Fanuc KAREL source: kt00308.KL

-- PROVISIONAL review KL for V1013-1; original PC SHA256 63806e7de99ed8727b65e89e63d5fef86488480187000dec51ab389faf893b3d
-- Incomplete behavior may be omitted. Consult companion uncertainty JSON. Do not deploy.
PROGRAM KT00308
%NOLOCKGROUP
VAR
  R2 : REAL
  OUT : BOOLEAN
-- UNRESOLVED_DECL H1 type=002017
BEGIN
  -- UNRESOLVED_PC offsets 5-19; opcodes 2E,22,9D,33,B4
  -- UNRESOLVED_PC offsets 24-35; opcodes 2E,23
  -- UNRESOLVED_PC offsets 40-64; opcodes 22,9D,33,B3,21,29,64,6E,23
  -- UNRESOLVED_PC offsets 69-73; opcodes 7F
END KT00308
